// TIA Portal V20 export
TYPE "AZ_Struct_PLC2Drv"
   STRUCT
      RemoteIO_IN : Word;
      OperNumSel : Word;
      FixedIO_IN { S7_SetPoint := 'True'} : "AZ_FixedIO_PLC2Drv";
      DDO_Type : Word;
      DDO_Pos : DInt;
      DDO_Vel : DInt;
      DDO_Acc : UDInt;
      DDO_Dec : UDInt;
      DDO_Crnt : UInt;
      DDO_Trans : Word;
      Reserve : Word;
      ReadPrmID : Word;
      WriteReq : Word;
      WritePrmID : Word;
      WriteData : DInt;
   END_STRUCT;
END_TYPE
